FUNCTION_BLOCK T_SafeTon_Tests EXTENDS TcUnit.FB_TestSuite
VAR
    // Test_OutputDelayedOn
    group_1 : T_SafeGroup;
    fb_1 : T_SafeTon(group := group_1) := (Parameters := (DelayTime := T#100MS));
    state_1 : INT := 10;
    waitTimer_1 : TON;
    // Test_UnconnectedInputIsRefused
    group_2 : T_SafeGroup;
    fb_2 : T_SafeTon(group := group_2);
END_VAR

Test_OutputDelayedOn();
Test_UnconnectedInputIsRefused();

METHOD PRIVATE Test_OutputDelayedOn
TcUnit.TEST(__POUNAME());
waitTimer_1();

CASE state_1 OF
    10:
        // act
        group_1(Run := TRUE);
        fb_1(TonIn1 := TRUE);
        // assert
        AssertEquals_BOOL(Expected := FALSE, Actual := fb_1.TonOut, Message := 'output not yet on');
        AssertEquals_BYTE(Expected := TO_BYTE(E_SafeTonState.DelayIn), Actual := fb_1.State, Message := 'state DELAYIN');
        state_1 := 20;
        waitTimer_1(IN := TRUE, PT := T#200MS);
    20:
        group_1(Run := TRUE);
        fb_1(TonIn1 := TRUE);

        IF NOT waitTimer_1.Q THEN
            RETURN;
        END_IF

        waitTimer_1(IN := FALSE);
        // assert
        AssertEquals_BOOL(Expected := TRUE, Actual := fb_1.TonOut, Message := 'output on after the delay');
        fb_1(TonIn1 := FALSE);
        AssertEquals_BOOL(Expected := FALSE, Actual := fb_1.TonOut, Message := 'output off immediately');
        TEST_FINISHED_NAMED(__POUNAME());
        state_1 := 10;
END_CASE
END_METHOD

METHOD PRIVATE Test_UnconnectedInputIsRefused
TcUnit.TEST(__POUNAME());
// arrange / act: TonIn1 is unconnected, which the Safety Editor refuses
group_2(Run := TRUE);
fb_2();
group_2(Run := TRUE);
fb_2();
// assert
AssertEquals_BOOL(Expected := TRUE, Actual := fb_2.Error, Message := 'configuration error reported');
AssertEquals_BYTE(Expected := TO_BYTE(E_SafeFbState.Error), Actual := fb_2.State, Message := 'state ERROR');
AssertEquals_WORD(Expected := WORD#16#8000, Actual := fb_2.Diag, Message := 'diag bit 15 configuration refused');
AssertEquals_BOOL(Expected := FALSE, Actual := fb_2.TonOut, Message := 'TonOut stays at its safe value');
AssertEquals_BOOL(Expected := TRUE, Actual := group_2.FbErr, Message := 'the group sees an FB error');
// act: ErrAck 0 -> 1 -> 0 does not clear a configuration error
group_2(Run := TRUE, ErrAck := TRUE);
fb_2();
group_2(Run := TRUE, ErrAck := TRUE);
fb_2();
group_2(Run := TRUE, ErrAck := FALSE);
fb_2();
AssertEquals_BOOL(Expected := TRUE, Actual := fb_2.Error, Message := 'error not acknowledged');
AssertEquals_WORD(Expected := WORD#16#8000, Actual := fb_2.Diag, Message := 'diag bit 15 kept');
TEST_FINISHED_NAMED(__POUNAME());
END_METHOD

END_FUNCTION_BLOCK

(* stored: Version 1.1.0.1
   POU T_SafeTon_Tests: Id {0246d7a3-1b43-5c52-9a5a-d537dc1999e0}, SpecialFunc None
   Method Test_OutputDelayedOn: Id {8c094113-831d-5f18-a4a7-ca612caea250}
   Method Test_UnconnectedInputIsRefused: Id {076d468e-d757-4e3d-aa66-a4c264c470d8} *)
